(* IEC 61131-3 sources: realtime-platform-1.0/plc-program, 3 files *)

(* ---- Bench_Main.st ---- *)
VAR
lastClock : BOOL;
sampleIdx : INT;
bufT0 : REAL;
bufT1 : REAL;
bufT2 : REAL;
bufT3 : REAL;
bufT4 : REAL;
bufT5 : REAL;
bufT6 : REAL;
bufT7 : REAL;
bufT8 : REAL;
bufT9 : REAL;
bufP0 : REAL;
bufP1 : REAL;
bufP2 : REAL;
bufP3 : REAL;
bufP4 : REAL;
bufP5 : REAL;
bufP6 : REAL;
bufP7 : REAL;
bufP8 : REAL;
bufP9 : REAL;
bufH0 : REAL;
bufH1 : REAL;
bufH2 : REAL;
bufH3 : REAL;
bufH4 : REAL;
bufH5 : REAL;
bufH6 : REAL;
bufH7 : REAL;
bufH8 : REAL;
bufH9 : REAL;
fifoSumT : REAL;
fifoSumP : REAL;
fifoSumH : REAL;
fifoAvgT : REAL;
fifoAvgP : REAL;
fifoAvgH : REAL;
abnormal : INT;
statusWord : INT;
aiTemp : REAL;
aiPress : REAL;
aiHumid : REAL;
raw4mA : REAL;
raw20mA : REAL;
rawSpan : REAL;
pressSet : REAL;
heightSet : REAL;
localMode : BOOL;
runFlag : BOOL;
x0Last : BOOL;
cycleStep : INT;
cycleCount : INT;
tickCnt : INT;
baseH : INT;
topH : INT;
upTicks : INT;
holdTicks : INT;
maxCycles : INT;
yUp : BOOL;
yDown : BOOL;
END_VAR

(************************************************************
 * Bench_Main.st —— 台架实测主程序（LiteST 兼容版）
 * 机型：汇川 Easy320（AutoShop，结构化文本 LiteST）
 *
 * ⚠️ 本版按 LiteST 限制改写：
 *   · 不用 ARRAY，不用 Arr[n] 下标（LiteST 不支持变量下标）
 *   · 不用 FOR 循环
 *   · 10 点滑窗改成 30 个标量移位寄存器（bufT0..bufT9 / bufP0..bufP9 / bufH0..bufH9）
 *
 * 功能：
 *   ① 协议：100 ms 采样、10 点均值、1 s 组包、状态字、序号、子包
 *   ② 本地循环：X0 启动、X1 停止、X2 常闭急停；20 s 升 / 60 s 顶保 /
 *      20 s 降 / 60 s 底保，30 次自动停；X3 选本地/远程
 *   ③ 安全：Y0/Y1 互锁；急停保持位置不降弓；D2022 钳位 50~1450
 *
 * 模式：
 *   X3 = 0  远程：D2021/D2022 由平台 FC16 写入
 *   X3 = 1  本地：PLC 自己写 D2022，按 100→1400→100 循环
 *
 * 寄存器：D2001 温度×10  D2002 压力×10  D2003 湿度×10
 *         D2004 状态字  D2005 序号  D2011-15 子包
 *         D2021 压力设定×10kPa  D2022 高度设定 mm
 *
 * 下载前替换 5 个软元件（按实际模块地址核对）：
 *   温度 D500  压力 D501  湿度 D502  比例阀 D510  升弓 D511（模块到位后换回 AIW/AQW）
 ************************************************************)

(* ============================================================
 * 每 100 ms 执行一次（M8012 上升沿）
 * ============================================================ *)
IF M8012 AND NOT lastClock THEN

    (* 常量每周期赋值，避免依赖变量初值 *)
    raw4mA := 8000.0;
    raw20mA := 40000.0;
    rawSpan := 32000.0;
    baseH := 100;
    topH := 1400;
    upTicks := 200;
    holdTicks := 600;
    maxCycles := 30;

    (* ---------- 1. 4~20 mA → 工程量 ---------- *)
    aiTemp  := (D500 - raw4mA) / rawSpan * 90.0 - 10.0;
    aiPress := (D501 - raw4mA) / rawSpan * 1000.0;
    aiHumid := (D502 - raw4mA) / rawSpan * 100.0;

    (* ---------- 2. 移位寄存器：新值进 bufT0，旧值后移 ---------- *)
    bufT9 := bufT8; bufT8 := bufT7; bufT7 := bufT6; bufT6 := bufT5; bufT5 := bufT4;
    bufT4 := bufT3; bufT3 := bufT2; bufT2 := bufT1; bufT1 := bufT0; bufT0 := aiTemp;

    bufP9 := bufP8; bufP8 := bufP7; bufP7 := bufP6; bufP6 := bufP5; bufP5 := bufP4;
    bufP4 := bufP3; bufP3 := bufP2; bufP2 := bufP1; bufP1 := bufP0; bufP0 := aiPress;

    bufH9 := bufH8; bufH8 := bufH7; bufH7 := bufH6; bufH6 := bufH5; bufH5 := bufH4;
    bufH4 := bufH3; bufH3 := bufH2; bufH2 := bufH1; bufH1 := bufH0; bufH0 := aiHumid;

    (* ---------- 3. 每 10 个采样（1 s）组包 ---------- *)
    sampleIdx := sampleIdx + 1;
    IF sampleIdx >= 10 THEN
        sampleIdx := 0;

        fifoSumT := bufT0+bufT1+bufT2+bufT3+bufT4+bufT5+bufT6+bufT7+bufT8+bufT9;
        fifoSumP := bufP0+bufP1+bufP2+bufP3+bufP4+bufP5+bufP6+bufP7+bufP8+bufP9;
        fifoSumH := bufH0+bufH1+bufH2+bufH3+bufH4+bufH5+bufH6+bufH7+bufH8+bufH9;
        fifoAvgT := fifoSumT / 10.0;
        fifoAvgP := fifoSumP / 10.0;
        fifoAvgH := fifoSumH / 10.0;

        (* ---------- 4. 阈值判定 ---------- *)
        abnormal := 0;
        IF fifoAvgT > 80.0 OR fifoAvgT < -10.0 THEN abnormal := abnormal OR 1;   END_IF;
        IF fifoAvgP > 1000.0 OR fifoAvgP < 100.0 THEN abnormal := abnormal OR 2; END_IF;
        IF fifoAvgH > 85.0 THEN abnormal := abnormal OR 4;                   END_IF;

        (* ---------- 5. 主包 ---------- *)
        D2001 := REAL_TO_INT(fifoAvgT * 10.0);
        IF fifoAvgT < 0.0 THEN D2001 := D2001 + 65536; END_IF;
        D2002 := REAL_TO_INT(fifoAvgP * 10.0);
        D2003 := REAL_TO_INT(fifoAvgH * 10.0);

        (* ---------- 6. 序号回绕 ---------- *)
        D2005 := D2005 + 1;
        IF D2005 > 65535 THEN D2005 := 1; END_IF;

        (* ---------- 7. 状态字 + 子包 ---------- *)
        statusWord := 16#40;
        IF abnormal <> 0 THEN
            statusWord := statusWord OR abnormal;
            statusWord := statusWord OR 16#80;
            D2011 := D2005;
            D2012 := abnormal;
            D2013 := D2001;
            D2014 := D2002;
            D2015 := D2003;
        END_IF;
        D2004 := statusWord;
    END_IF;

    (* ---------- 8. 设定值安全钳位 ---------- *)
    IF D2022 < 50 THEN D2022 := 50; END_IF;
    IF D2022 > 1450 THEN D2022 := 1450; END_IF;
    IF D2021 < 0 THEN D2021 := 0; END_IF;
    IF D2021 > 10000 THEN D2021 := 10000; END_IF;

    (* ---------- 9. 本地循环（X3=1） ---------- *)
    localMode := X3;
    IF NOT localMode THEN
        runFlag := FALSE;
        cycleStep := 0;
        tickCnt := 0;
        yUp := FALSE;
        yDown := FALSE;
    ELSE
        (* 急停/停止：X2 常闭（正常=1，按下=0）；X1 常开（按下=1） *)
        IF (NOT X2) OR X1 THEN
            runFlag := FALSE;
            cycleStep := 0;
            tickCnt := 0;
            yUp := FALSE;
            yDown := FALSE;
        END_IF;

        (* 启动：X0 上升沿 *)
        IF X0 AND NOT x0Last THEN
            runFlag := TRUE;
            cycleCount := 0;
            cycleStep := 1;
            tickCnt := 0;
        END_IF;

        IF runFlag THEN
            tickCnt := tickCnt + 1;
            IF cycleStep = 1 THEN
                yUp := TRUE; yDown := FALSE; D2022 := topH;
                IF tickCnt >= upTicks THEN
                    cycleStep := 2; tickCnt := 0; yUp := FALSE;
                END_IF;
            ELSIF cycleStep = 2 THEN
                yUp := FALSE; yDown := FALSE; D2022 := topH;
                IF tickCnt >= holdTicks THEN
                    cycleStep := 3; tickCnt := 0;
                END_IF;
            ELSIF cycleStep = 3 THEN
                yUp := FALSE; yDown := TRUE; D2022 := baseH;
                IF tickCnt >= upTicks THEN
                    cycleStep := 4; tickCnt := 0; yDown := FALSE;
                END_IF;
            ELSIF cycleStep = 4 THEN
                yUp := FALSE; yDown := FALSE; D2022 := baseH;
                IF tickCnt >= holdTicks THEN
                    cycleCount := cycleCount + 1;
                    tickCnt := 0;
                    IF cycleCount >= maxCycles THEN
                        runFlag := FALSE;
                        cycleStep := 0;
                        D2022 := baseH;
                    ELSE
                        cycleStep := 1;
                    END_IF;
                END_IF;
            END_IF;
        END_IF;
        (* 急停/停止保持当前位置，不主动降弓 *)
    END_IF;

    (* X0 边沿记忆每周期更新 *)
    x0Last := X0;

    (* ---------- 10. 输出互锁 ---------- *)
    IF yUp AND yDown THEN
        yUp := FALSE;
        yDown := FALSE;
    END_IF;
    Y0 := yUp;
    Y1 := yDown;

    (* ---------- 11. AO 输出（按全行程 1500 mm 标定） ---------- *)
    pressSet  := D2021 / 10.0;
    heightSet := D2022;
    D510   := REAL_TO_INT((pressSet  / 1000.0) * rawSpan + raw4mA);
    D511 := REAL_TO_INT((heightSet / 1500.0) * rawSpan + raw4mA);

END_IF;

lastClock := M8012;

(* 下载前检查：
   1) 5 个软元件替换为实际地址；
   2) MBS 从站 502、unit 1，4xN ↔ DN 映射；
   3) X3=0 远程 / X3=1 本地；X2 必须接常闭急停。 *)

(* ---- Bench_Main_noVAR.st ---- *)
(************************************************************
 * Bench_Main.st —— 台架实测主程序（LiteST 兼容版）
 * 机型：汇川 Easy320（AutoShop，结构化文本 LiteST）
 *
 * ⚠️ 本版按 LiteST 限制改写：
 *   · 不用 ARRAY，不用 Arr[n] 下标（LiteST 不支持变量下标）
 *   · 不用 FOR 循环
 *   · 10 点滑窗改成 30 个标量移位寄存器（bufT0..bufT9 / bufP0..bufP9 / bufH0..bufH9）
 *
 * 功能：
 *   ① 协议：100 ms 采样、10 点均值、1 s 组包、状态字、序号、子包
 *   ② 本地循环：X0 启动、X1 停止、X2 常闭急停；20 s 升 / 60 s 顶保 /
 *      20 s 降 / 60 s 底保，30 次自动停；X3 选本地/远程
 *   ③ 安全：Y0/Y1 互锁；急停保持位置不降弓；D2022 钳位 50~1450
 *
 * 模式：
 *   X3 = 0  远程：D2021/D2022 由平台 FC16 写入
 *   X3 = 1  本地：PLC 自己写 D2022，按 100→1400→100 循环
 *
 * 寄存器：D2001 温度×10  D2002 压力×10  D2003 湿度×10
 *         D2004 状态字  D2005 序号  D2011-15 子包
 *         D2021 压力设定×10kPa  D2022 高度设定 mm
 *
 * 下载前替换 5 个软元件（按实际模块地址核对）：
 *   温度 D500  压力 D501  湿度 D502  比例阀 D510  升弓 D511（模块到位后换回 AIW/AQW）
 ************************************************************)

(* ============================================================
 * 每 100 ms 执行一次（M8012 上升沿）
 * ============================================================ *)
IF M8012 AND NOT lastClock THEN

    (* 常量每周期赋值，避免依赖变量初值 *)
    raw4mA := 8000.0;
    raw20mA := 40000.0;
    rawSpan := 32000.0;
    baseH := 100;
    topH := 1400;
    upTicks := 200;
    holdTicks := 600;
    maxCycles := 30;

    (* ---------- 1. 4~20 mA → 工程量 ---------- *)
    aiTemp  := (D500 - raw4mA) / rawSpan * 90.0 - 10.0;
    aiPress := (D501 - raw4mA) / rawSpan * 1000.0;
    aiHumid := (D502 - raw4mA) / rawSpan * 100.0;

    (* ---------- 2. 移位寄存器：新值进 bufT0，旧值后移 ---------- *)
    bufT9 := bufT8; bufT8 := bufT7; bufT7 := bufT6; bufT6 := bufT5; bufT5 := bufT4;
    bufT4 := bufT3; bufT3 := bufT2; bufT2 := bufT1; bufT1 := bufT0; bufT0 := aiTemp;

    bufP9 := bufP8; bufP8 := bufP7; bufP7 := bufP6; bufP6 := bufP5; bufP5 := bufP4;
    bufP4 := bufP3; bufP3 := bufP2; bufP2 := bufP1; bufP1 := bufP0; bufP0 := aiPress;

    bufH9 := bufH8; bufH8 := bufH7; bufH7 := bufH6; bufH6 := bufH5; bufH5 := bufH4;
    bufH4 := bufH3; bufH3 := bufH2; bufH2 := bufH1; bufH1 := bufH0; bufH0 := aiHumid;

    (* ---------- 3. 每 10 个采样（1 s）组包 ---------- *)
    sampleIdx := sampleIdx + 1;
    IF sampleIdx >= 10 THEN
        sampleIdx := 0;

        fifoSumT := bufT0+bufT1+bufT2+bufT3+bufT4+bufT5+bufT6+bufT7+bufT8+bufT9;
        fifoSumP := bufP0+bufP1+bufP2+bufP3+bufP4+bufP5+bufP6+bufP7+bufP8+bufP9;
        fifoSumH := bufH0+bufH1+bufH2+bufH3+bufH4+bufH5+bufH6+bufH7+bufH8+bufH9;
        fifoAvgT := fifoSumT / 10.0;
        fifoAvgP := fifoSumP / 10.0;
        fifoAvgH := fifoSumH / 10.0;

        (* ---------- 4. 阈值判定 ---------- *)
        abnormal := 0;
        IF fifoAvgT > 80.0 OR fifoAvgT < -10.0 THEN abnormal := abnormal OR 1;   END_IF;
        IF fifoAvgP > 1000.0 OR fifoAvgP < 100.0 THEN abnormal := abnormal OR 2; END_IF;
        IF fifoAvgH > 85.0 THEN abnormal := abnormal OR 4;                   END_IF;

        (* ---------- 5. 主包 ---------- *)
        D2001 := REAL_TO_INT(fifoAvgT * 10.0);
        IF fifoAvgT < 0.0 THEN D2001 := D2001 + 65536; END_IF;
        D2002 := REAL_TO_INT(fifoAvgP * 10.0);
        D2003 := REAL_TO_INT(fifoAvgH * 10.0);

        (* ---------- 6. 序号回绕 ---------- *)
        D2005 := D2005 + 1;
        IF D2005 > 65535 THEN D2005 := 1; END_IF;

        (* ---------- 7. 状态字 + 子包 ---------- *)
        statusWord := 16#40;
        IF abnormal <> 0 THEN
            statusWord := statusWord OR abnormal;
            statusWord := statusWord OR 16#80;
            D2011 := D2005;
            D2012 := abnormal;
            D2013 := D2001;
            D2014 := D2002;
            D2015 := D2003;
        END_IF;
        D2004 := statusWord;
    END_IF;

    (* ---------- 8. 设定值安全钳位 ---------- *)
    IF D2022 < 50 THEN D2022 := 50; END_IF;
    IF D2022 > 1450 THEN D2022 := 1450; END_IF;
    IF D2021 < 0 THEN D2021 := 0; END_IF;
    IF D2021 > 10000 THEN D2021 := 10000; END_IF;

    (* ---------- 9. 本地循环（X3=1） ---------- *)
    localMode := X3;
    IF NOT localMode THEN
        runFlag := FALSE;
        cycleStep := 0;
        tickCnt := 0;
        yUp := FALSE;
        yDown := FALSE;
    ELSE
        (* 急停/停止：X2 常闭（正常=1，按下=0）；X1 常开（按下=1） *)
        IF (NOT X2) OR X1 THEN
            runFlag := FALSE;
            cycleStep := 0;
            tickCnt := 0;
            yUp := FALSE;
            yDown := FALSE;
        END_IF;

        (* 启动：X0 上升沿 *)
        IF X0 AND NOT x0Last THEN
            runFlag := TRUE;
            cycleCount := 0;
            cycleStep := 1;
            tickCnt := 0;
        END_IF;

        IF runFlag THEN
            tickCnt := tickCnt + 1;
            IF cycleStep = 1 THEN
                yUp := TRUE; yDown := FALSE; D2022 := topH;
                IF tickCnt >= upTicks THEN
                    cycleStep := 2; tickCnt := 0; yUp := FALSE;
                END_IF;
            ELSIF cycleStep = 2 THEN
                yUp := FALSE; yDown := FALSE; D2022 := topH;
                IF tickCnt >= holdTicks THEN
                    cycleStep := 3; tickCnt := 0;
                END_IF;
            ELSIF cycleStep = 3 THEN
                yUp := FALSE; yDown := TRUE; D2022 := baseH;
                IF tickCnt >= upTicks THEN
                    cycleStep := 4; tickCnt := 0; yDown := FALSE;
                END_IF;
            ELSIF cycleStep = 4 THEN
                yUp := FALSE; yDown := FALSE; D2022 := baseH;
                IF tickCnt >= holdTicks THEN
                    cycleCount := cycleCount + 1;
                    tickCnt := 0;
                    IF cycleCount >= maxCycles THEN
                        runFlag := FALSE;
                        cycleStep := 0;
                        D2022 := baseH;
                    ELSE
                        cycleStep := 1;
                    END_IF;
                END_IF;
            END_IF;
        END_IF;
        (* 急停/停止保持当前位置，不主动降弓 *)
    END_IF;

    (* X0 边沿记忆每周期更新 *)
    x0Last := X0;

    (* ---------- 10. 输出互锁 ---------- *)
    IF yUp AND yDown THEN
        yUp := FALSE;
        yDown := FALSE;
    END_IF;
    Y0 := yUp;
    Y1 := yDown;

    (* ---------- 11. AO 输出（按全行程 1500 mm 标定） ---------- *)
    pressSet  := D2021 / 10.0;
    heightSet := D2022;
    D510   := REAL_TO_INT((pressSet  / 1000.0) * rawSpan + raw4mA);
    D511 := REAL_TO_INT((heightSet / 1500.0) * rawSpan + raw4mA);

END_IF;

lastClock := M8012;

(* 下载前检查：
   1) 5 个软元件替换为实际地址；
   2) MBS 从站 502、unit 1，4xN ↔ DN 映射；
   3) X3=0 远程 / X3=1 本地；X2 必须接常闭急停。 *)

(* ---- Easy320_main.st ---- *)
(************************************************************
 * Easy320_main.st —— 汇川 Easy320 传感器采集 + Modbus 组包参考程序
 * 语言: ST（AutoShop 编译下载）  目标: 文档级参考代码
 *
 * 功能: 100ms 采样温度/压力/湿度(4-20mA) → 10 条滑窗均值
 *       → 阈值判异常 → 主包(全部数据) + 子包(异常数据)
 *       → 状态字/序号 → 读回写寄存器驱动比例阀/升弓机构
 *
 * 机型: 汇川 Easy320（Easy 系列紧凑型网络主机，双网口，AutoShop 编程）
 * ⚠️ D 区 ↔ Modbus 映射（AutoShop MBS 服务: 4xN ↔ DN 直接对应）
 *    本程序用 D2001-D2022。Easy320 属 Easy 系列，D 区从 D0 起编址，
 *    没有 D30001 段（该段只存在于 D 区容量 ≥32767 的大容量机型）。
 *    平台 .env 默认值已与之一致（协议地址 = 这里选定的 4x 地址）：
 *        PLC_REG_TEMP=2001  PLC_REG_PRESS=2002  PLC_REG_HUMID=2003
 *        PLC_REG_STATUS=2004  PLC_REG_SEQ=2005
 *        PLC_REG_SUB_BASE=2011  PLC_REG_WRITE_FORCE=2021  PLC_REG_WRITE_HEIGHT=2022
 *    仅在换用 D 区 ≥32767 的大容量机型时，才把 D2001-2022 整体替换为
 *    D30001-30022 段，并同步把平台 .env 的 PLC_REG_* 改到 30001 起。
 *
 * 寄存器语义（协议原地址 = 4x + 本程序 D 编号）：
 *   D2001     温度均值 ×10（有符号 16 位，负数用补码）
 *   D2002     压力均值 ×10（0.1kPa，勿用 ×100：1000kPa→100000 超 uint16）
 *   D2003     湿度均值 ×10
 *   D2004     状态字 bit0/1/2=温/压/湿异常；bit6=0x40 扩展协议标志(恒置)；
 *             bit7=0x80 子包有效
 *   D2005     主包序号（65535→1 回绕，0 保留给旧固件）
 *   D2011     子包序号（= 异常发生时主包序号）
 *   D2012     异常位图（bit0-2 同状态字）
 *   D2013-15  子包异常值（温度/压力/湿度，缩放同上，仅对应位有效）
 *   D2021     接触力环输出 = 气囊压力设定 ×10 kPa   [平台 FC16 写入]
 *   D2022     姿态环输出   = 弓头高度设定 mm         [平台 FC16 写入]
 ************************************************************)

VAR
    (* ---- 采样与滑窗 ---- *)
    lastClock   : BOOL;                     (* 100ms 脉冲上升沿检测 *)
    sampleIdx   : INT := 0;                 (* 当前滑窗位置 0-9 *)
    fifoT       : ARRAY[0..9] OF REAL;      (* 温度滑窗 FIFO *)
    fifoP       : ARRAY[0..9] OF REAL;      (* 压力滑窗 FIFO *)
    fifoH       : ARRAY[0..9] OF REAL;      (* 湿度滑窗 FIFO *)
    sumT, sumP, sumH : REAL;                (* 滑窗求和 *)
    avgT, avgP, avgH : REAL;                (* 10 条均值 *)
    i           : INT;                      (* 循环变量 *)

    (* ---- 阈值判定 ---- *)
    abnormal    : INT := 0;                 (* 异常位图 0=正常 bit0温 bit1压 bit2湿 *)
    statusWord  : INT := 0;                 (* D2004 状态字组装用 *)

    (* ---- 模拟量原始值（请替换为实际 AD 通道元件）---- *)
    aiTemp      : REAL;                     (* 温度通道原始值 *)
    aiPress     : REAL;                     (* 压力通道原始值 *)
    aiHumid     : REAL;                     (* 湿度通道原始值 *)

    (* ---- 模拟量量程（GL10-4AD: 4mA/20mA 对应原始值，按实际模块校准）---- *)
    raw4mA      : REAL := 8000.0;
    raw20mA     : REAL := 40000.0;
    rawSpan     : REAL := 32000.0;          (* raw20mA - raw4mA *)

    (* ---- 写回读值 ---- *)
    pressSet    : REAL;                     (* 来自 D2021 的压力设定 kPa *)
    heightSet   : REAL;                     (* 来自 D2022 的高度设定 mm *)
END_VAR

(* ============================================================
 * 主流程：每 100ms 执行一次（AutoShop 的 100ms 脉冲继电器 SM4010；
 * Easy320 沿用同一套特殊软元件编号，若你的机型手册中该位不同，请替换）
 * ============================================================ *)
IF SM4010 AND NOT lastClock THEN

    (* ---------- 1. 4-20mA → 工程量换算（量程按实际传感器标定修改） ----------
       温度: 4-20mA 对应 -10 ~ 80°C
       压力: 4-20mA 对应   0 ~ 1000kPa
       湿度: 4-20mA 对应   0 ~ 100%RH                            *)
    aiTemp  := (温度通道元件 - raw4mA) / rawSpan * 90.0 - 10.0;
    aiPress := (压力通道元件 - raw4mA) / rawSpan * 1000.0;
    aiHumid := (湿度通道元件 - raw4mA) / rawSpan * 100.0;

    (* ---------- 2. 滑窗 FIFO：新样本覆盖最旧的一条 ---------- *)
    fifoT[sampleIdx] := aiTemp;
    fifoP[sampleIdx] := aiPress;
    fifoH[sampleIdx] := aiHumid;
    sampleIdx := sampleIdx + 1;

    (* ---------- 3. 每满 10 条（1s）计算均值 + 判阈 + 组包 ---------- *)
    IF sampleIdx >= 10 THEN
        sampleIdx := 0;
        sumT := 0.0; sumP := 0.0; sumH := 0.0;
        FOR i := 0 TO 9 DO
            sumT := sumT + fifoT[i];
            sumP := sumP + fifoP[i];
            sumH := sumH + fifoH[i];
        END_FOR;
        avgT := sumT / 10.0;
        avgP := sumP / 10.0;
        avgH := sumH / 10.0;

        (* ---------- 4. 阈值判定（与平台 THRESHOLDS 保持一致） ---------- *)
        abnormal := 0;
        IF avgT > 80.0 OR avgT < -10.0 THEN abnormal := abnormal OR 1;   END_IF;
        IF avgP > 1000.0 OR avgP < 100.0 THEN abnormal := abnormal OR 2; END_IF;
        IF avgH > 85.0 THEN abnormal := abnormal OR 4;                   END_IF;

        (* ---------- 5. 主包写入（全部数据） ----------
           REAL→定点：四舍五入到 0.1 精度；温度负值补码处理         *)
        D2001 := REAL_TO_INT(avgT * 10.0);                  (* 温度 ×10 *)
        IF avgT < 0.0 THEN D2001 := D2001 + 65536; END_IF;  (* 负数补码 *)
        D2002 := REAL_TO_INT(avgP * 10.0);                  (* 压力 ×10 *)
        D2003 := REAL_TO_INT(avgH * 10.0);                  (* 湿度 ×10 *)

        (* ---------- 6. 序号：65535→1 回绕（0 保留给旧固件判定） ---------- *)
        D2005 := D2005 + 1;
        IF D2005 > 65535 THEN D2005 := 1; END_IF;

        (* ---------- 7. 状态字：bit6 恒置扩展协议标志；异常时置对应位 ---------- *)
        statusWord := 16#40;                               (* bit6 恒置 *)
        IF abnormal <> 0 THEN
            statusWord := statusWord OR abnormal;          (* bit0-2 异常位 *)
            statusWord := statusWord OR 16#80;             (* bit7 子包有效 *)

            (* ---------- 8. 子包：序号=主包序号，位图+异常值 ---------- *)
            D2011 := D2005;
            D2012 := abnormal;
            D2013 := D2001;                                (* 异常值 = 本周期均值 *)
            D2014 := D2002;
            D2015 := D2003;
        END_IF;
        D2004 := statusWord;

        (* ---------- 9. 读回平台写寄存器，驱动执行机构 ----------
           D2021 压力设定(×10 kPa) → 比例阀模拟量输出
           D2022 高度设定(mm)     → 升弓机构模拟量输出
           （量程换算按实际执行机构标定修改）                     *)
        pressSet  := D2021 / 10.0;                         (* kPa *)
        heightSet := D2022;                                (* mm *)
        比例阀输出元件 := REAL_TO_INT((pressSet  / 1000.0) * rawSpan + raw4mA);
        升弓机构输出元件 := REAL_TO_INT((heightSet / 2600.0) * rawSpan + raw4mA);
    END_IF;
END_IF;

lastClock := SM4010;

(* 程序结束。下载到 PLC 前请务必：
   1) 替换"温度通道元件/压力通道元件/湿度通道元件/比例阀输出元件/升弓机构输出元件"
      为实际软元件；
   2) 在 MBS 服务配置中启用从站（端口 502）并确认 4xN ↔ DN 映射；
   3) 用 ModbusPoll 读 4x2001-2005 核对数值与状态字（bit6=0x40）；
   4) 平台 .env 按本文件头部的映射表设置 REG_* 变量。 *)
